(* IEC 61131-3 sources: llm-plc-st-eval/data/processed_v2/gpt-4o/I6/zero_shot, 3 files *)

(* ---- ejec_1.st ---- *)
FUNCTION_BLOCK FB_Temperatura
VAR_INPUT
    rawTemp : INT; // Valor de entrada de la temperatura en formato entero
END_VAR

VAR_OUTPUT
    tempC : REAL; // Temperatura calculada en grados Celsius
    enfriador : BOOL; // Estado del enfriador
    almSensor : BOOL; // Alarma de sensor
END_VAR

VAR
    tempC_prev : REAL; // Valor previo de la temperatura en grados Celsius
END_VAR

// Conversión del valor de entrada a grados Celsius
tempC := (REAL(rawTemp) * 100.0) / 27648.0;

// Verificación de los límites del sensor
IF (rawTemp < 0) OR (rawTemp > 27648) THEN
    almSensor := TRUE; // Activar alarma de sensor
    enfriador := FALSE; // Desactivar enfriador
ELSE
    almSensor := FALSE; // Desactivar alarma de sensor

    // Control del enfriador con histéresis
    IF tempC >= 80.0 THEN
        enfriador := TRUE; // Activar enfriador
    ELSIF tempC <= 75.0 THEN
        enfriador := FALSE; // Desactivar enfriador
    ELSE
        // Mantener el estado actual del enfriador
        enfriador := enfriador;
    END_IF
END_IF
END_FUNCTION_BLOCK

(* ---- ejec_2.st ---- *)
FUNCTION_BLOCK FB_Temperatura
VAR_INPUT
    rawTemp : INT; // Valor de entrada de temperatura en bruto
END_VAR

VAR_OUTPUT
    tempC : REAL; // Temperatura calculada en grados Celsius
    enfriador : BOOL; // Estado del enfriador
    almSensor : BOOL; // Alarma de sensor
END_VAR

VAR
    tempC_prev : REAL; // Temperatura anterior para control de histéresis
END_VAR

// Conversión de rawTemp a grados Celsius
tempC := (REAL(rawTemp) * 100.0) / 27648.0;

// Comprobación de límites de rawTemp para activar alarma
IF (rawTemp < 0) OR (rawTemp > 27648) THEN
    almSensor := TRUE;
    enfriador := FALSE; // Desactiva el enfriador si hay un error de sensor
ELSE
    almSensor := FALSE;

    // Control de histéresis para el enfriador
    IF tempC >= 80.0 THEN
        enfriador := TRUE;
    ELSIF tempC <= 75.0 THEN
        enfriador := FALSE;
    ELSE
        // Mantiene el estado anterior del enfriador
        enfriador := enfriador;
    END_IF;
END_IF;
END_FUNCTION_BLOCK

(* ---- ejec_3.st ---- *)
FUNCTION_BLOCK FB_Temperatura
VAR_INPUT
    rawTemp : INT; // Entrada de temperatura en bruto
END_VAR_INPUT

VAR_OUTPUT
    tempC : REAL; // Temperatura calculada en grados Celsius
    enfriador : BOOL; // Estado del enfriador
    almSensor : BOOL; // Alarma de sensor
END_VAR_OUTPUT

VAR
    tempC_prev : REAL; // Temperatura previa para control de histéresis
END_VAR

// Conversión de rawTemp a grados Celsius
tempC := (REAL(rawTemp) * 100.0) / 27648.0;

// Verificación de límites de rawTemp para activar alarma de sensor
IF (rawTemp < 0) OR (rawTemp > 27648) THEN
    almSensor := TRUE;
    enfriador := FALSE; // Desactiva el enfriador si hay error en el sensor
ELSE
    almSensor := FALSE;

    // Control del enfriador con histéresis
    IF tempC >= 80.0 THEN
        enfriador := TRUE;
    ELSIF tempC <= 75.0 THEN
        enfriador := FALSE;
    ELSE
        // Mantiene el estado anterior del enfriador
        enfriador := enfriador;
    END_IF;
END_IF;

END_FUNCTION_BLOCK
